PROGRAM PB_UnitTests
VAR
	TestRunner : T_TestRunner;
	
	Test1 : T_Test1;
	Test2 : T_Test2;
	Test3 : T_Test3;
	
	Init : BOOL := TRUE;
	
END_VAR

IF Init THEN
	Init := FALSE;
	TestRunner.ClearTests();
	TestRunner.AddTest(Test1);
	TestRunner.AddTest(Test2);
	TestRunner.AddTest(Test3);
END_IF

TestRunner.CyclicUpdate();

END_PROGRAM

(* stored: Version 1.1.0.1, ProductVersion 3.1.4024.15
   POU PB_UnitTests: Id {11d29a6e-06e7-4cc4-9e24-38d314218fa7}, SpecialFunc None *)
